(* IEC 61131-3 sources: llm-plc-st-eval/data/processed_definitivo/gemini-3.1-pro-preview/C7/zero_shot, 3 files *)

(* ---- ejec_1.st ---- *)
FUNCTION_BLOCK FB_Contador
VAR_INPUT
    sensorPieza : BOOL; // Contacto NA que alimenta la entrada de conteo
    btnReset : BOOL;    // Contacto NA que alimenta el reset del contador
END_VAR

VAR_OUTPUT
    loteListo : BOOL;   // Bobina que indica si se alcanzó el valor preestablecido
    cuenta : INT;       // Valor actual del contador
END_VAR

VAR
    C1 : CTU;           // Instancia del contador ascendente estándar
END_VAR

// Rama 1: Llamada al contador ascendente con límite de 12
C1(CU := sensorPieza, RESET := btnReset, PV := 12);

// Rama 2: Activación de la bobina loteListo con la salida Q del contador
loteListo := C1.Q;

// Rama 3: Transferencia del valor actual del contador a la salida cuenta
cuenta := C1.CV;

END_FUNCTION_BLOCK

(* ---- ejec_2.st ---- *)
FUNCTION_BLOCK FB_Contador
VAR_INPUT
    sensorPieza : BOOL; // Señal para incrementar el contador
    btnReset : BOOL;    // Señal para reiniciar el contador
END_VAR

VAR_OUTPUT
    loteListo : BOOL;   // Se activa al alcanzar el valor preestablecido
    cuenta : INT;       // Valor actual del conteo
END_VAR

VAR
    C1 : CTU;           // Instancia del contador ascendente
END_VAR

// Rama 1: Actualización del contador ascendente con PV = 12
C1(CU := sensorPieza, RESET := btnReset, PV := 12);

// Rama 2: La salida Q del contador activa la bobina loteListo
loteListo := C1.Q;

// Rama 3: Se transfiere el valor actual del contador a la salida cuenta
cuenta := C1.CV;

END_FUNCTION_BLOCK

(* ---- ejec_3.st ---- *)
FUNCTION_BLOCK FB_Contador
VAR_INPUT
    sensorPieza : BOOL; // Contacto normalmente abierto para conteo
    btnReset    : BOOL; // Contacto normalmente abierto para reinicio
END_VAR

VAR_OUTPUT
    loteListo   : BOOL; // Bobina que indica si el lote está completo
    cuenta      : INT;  // Valor actual del conteo
END_VAR

VAR
    C1          : CTU;  // Instancia del contador ascendente
END_VAR

// Rama 1: Actualización del contador ascendente con PV = 12
C1(
    CU := sensorPieza,
    RESET := btnReset,
    PV := 12
);

// Rama 2: La salida Q del contador activa la bobina loteListo
loteListo := C1.Q;

// Rama 3: Se transfiere el valor actual del contador a la variable cuenta
cuenta := C1.CV;

END_FUNCTION_BLOCK
